// TIA Portal V21 export
TagTable "T_V5"
  X_V5 :   (PLC tag Current_state_of_Bay0.Bay0[0,0], HMI_Connection_1, 100 ms)
